FUNCTION_BLOCK PID_FLAG_STATE_ACCESS (* Experimental read-only state interface; original PID arithmetic unchanged; native validation pending *)
  (* Standard: 61499-2 *)
  (* Version 0.1, 2026-10-20, Guilherme *)
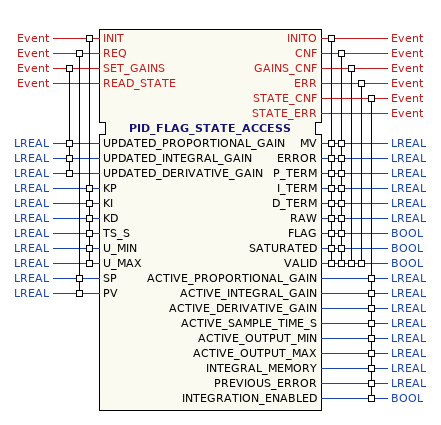
  EVENT_INPUT
    INIT WITH KP, KI, KD, TS_S, U_MIN, U_MAX;
    REQ WITH SP, PV;
    SET_GAINS WITH UPDATED_PROPORTIONAL_GAIN, UPDATED_INTEGRAL_GAIN, UPDATED_DERIVATIVE_GAIN;
    READ_STATE;
  END_EVENT
  EVENT_OUTPUT
    INITO WITH MV, ERROR, P_TERM, I_TERM, D_TERM, RAW, FLAG, SATURATED, VALID;
    CNF WITH MV, ERROR, P_TERM, I_TERM, D_TERM, RAW, FLAG, SATURATED, VALID;
    GAINS_CNF WITH VALID;
    ERR WITH VALID;
    STATE_CNF WITH ACTIVE_PROPORTIONAL_GAIN, ACTIVE_INTEGRAL_GAIN, ACTIVE_DERIVATIVE_GAIN, ACTIVE_SAMPLE_TIME_S, ACTIVE_OUTPUT_MIN, ACTIVE_OUTPUT_MAX, INTEGRAL_MEMORY, PREVIOUS_ERROR, INTEGRATION_ENABLED;
    STATE_ERR;
  END_EVENT
  VAR_INPUT
    UPDATED_PROPORTIONAL_GAIN : LREAL;
    UPDATED_INTEGRAL_GAIN : LREAL;
    UPDATED_DERIVATIVE_GAIN : LREAL;
    KP : LREAL;
    KI : LREAL;
    KD : LREAL;
    TS_S : LREAL;
    U_MIN : LREAL;
    U_MAX : LREAL;
    SP : LREAL;
    PV : LREAL;
  END_VAR
  VAR_OUTPUT
    MV : LREAL;
    ERROR : LREAL;
    P_TERM : LREAL;
    I_TERM : LREAL;
    D_TERM : LREAL;
    RAW : LREAL;
    FLAG : BOOL;
    SATURATED : BOOL;
    VALID : BOOL;
    ACTIVE_PROPORTIONAL_GAIN : LREAL;
    ACTIVE_INTEGRAL_GAIN : LREAL;
    ACTIVE_DERIVATIVE_GAIN : LREAL;
    ACTIVE_SAMPLE_TIME_S : LREAL;
    ACTIVE_OUTPUT_MIN : LREAL;
    ACTIVE_OUTPUT_MAX : LREAL;
    INTEGRAL_MEMORY : LREAL;
    PREVIOUS_ERROR : LREAL;
    INTEGRATION_ENABLED : BOOL;
  END_VAR
  VAR
    KP_ACTIVE : LREAL;
    KI_ACTIVE : LREAL;
    KD_ACTIVE : LREAL;
    TS_ACTIVE : LREAL;
    LOW : LREAL;
    HIGH : LREAL;
    I_MEMORY : LREAL;
    E_PREV : LREAL;
    E_NEXT : LREAL;
    I_NEXT : LREAL;
    D_NEXT : LREAL;
    P_NEXT : LREAL;
    IT_NEXT : LREAL;
    DT_NEXT : LREAL;
    RAW_NEXT : LREAL;
  END_VAR
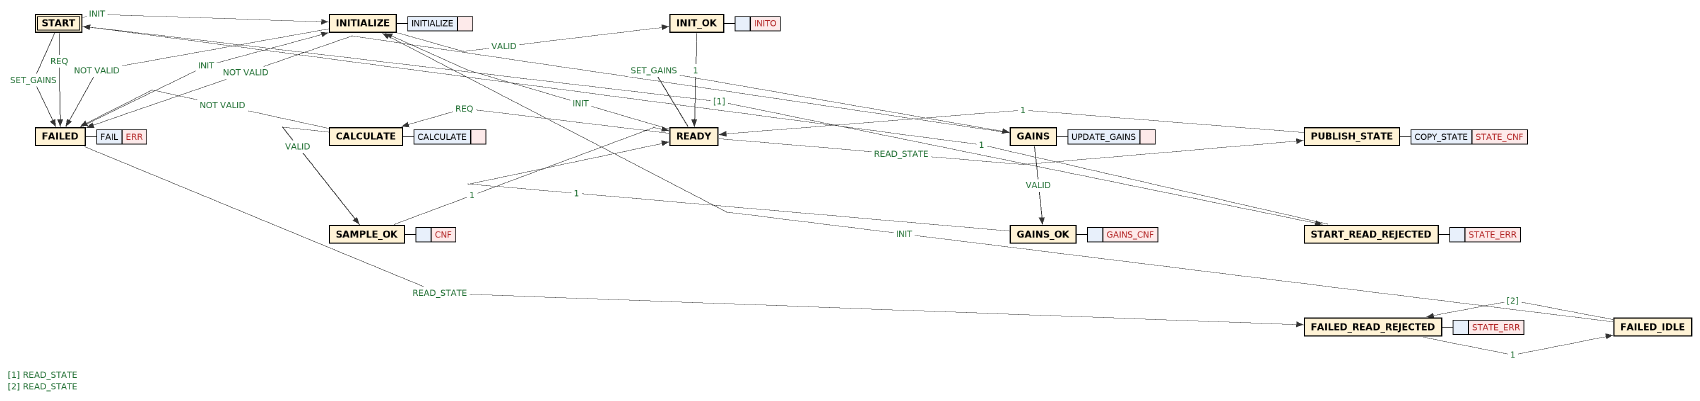
  EC_STATES
    START;
    FAILED_READ_REJECTED : -> STATE_ERR;
    START_READ_REJECTED : -> STATE_ERR;
    PUBLISH_STATE : COPY_STATE -> STATE_CNF;
    INITIALIZE : INITIALIZE;
    INIT_OK : -> INITO;
    READY;
    CALCULATE : CALCULATE;
    SAMPLE_OK : -> CNF;
    GAINS : UPDATE_GAINS;
    GAINS_OK : -> GAINS_CNF;
    FAILED : FAIL -> ERR;
    FAILED_IDLE;
  END_STATES
  EC_TRANSITIONS
    START TO INITIALIZE := INIT;
    START TO FAILED := REQ;
    START TO FAILED := SET_GAINS;
    INITIALIZE TO INIT_OK := VALID;
    INITIALIZE TO FAILED := NOT VALID;
    INIT_OK TO READY := 1;
    READY TO INITIALIZE := INIT;
    READY TO GAINS := SET_GAINS;
    READY TO CALCULATE := REQ;
    CALCULATE TO SAMPLE_OK := VALID;
    CALCULATE TO FAILED := NOT VALID;
    SAMPLE_OK TO READY := 1;
    GAINS TO GAINS_OK := VALID;
    GAINS TO FAILED := NOT VALID;
    GAINS_OK TO READY := 1;
    FAILED TO INITIALIZE := INIT;
    START TO START_READ_REJECTED := READ_STATE;
    START_READ_REJECTED TO START := 1;
    FAILED TO FAILED_READ_REJECTED := READ_STATE;
    FAILED_READ_REJECTED TO FAILED_IDLE := 1;
    FAILED_IDLE TO INITIALIZE := INIT;
    FAILED_IDLE TO FAILED_READ_REJECTED := READ_STATE;
    READY TO PUBLISH_STATE := READ_STATE;
    PUBLISH_STATE TO READY := 1;
  END_TRANSITIONS
  ALGORITHM INITIALIZE IN ST:
VALID := (KP >= -1.0E+100) AND (KP <= 1.0E+100) AND (KI >= -1.0E+100) AND (KI <= 1.0E+100) AND (KD >= -1.0E+100) AND (KD <= 1.0E+100) AND (TS_S >= -1.0E+100) AND (TS_S <= 1.0E+100) AND (U_MIN >= -1.0E+100) AND (U_MIN <= 1.0E+100) AND (U_MAX >= -1.0E+100) AND (U_MAX <= 1.0E+100) AND (TS_S > 0.0) AND (U_MIN < U_MAX);
IF VALID THEN
    KP_ACTIVE := KP;
    KI_ACTIVE := KI;
    KD_ACTIVE := KD;
    TS_ACTIVE := TS_S;
    LOW := U_MIN;
    HIGH := U_MAX;
    I_MEMORY := 0.0;
    E_PREV := 0.0;
    FLAG := TRUE;
    MV := 0.0;
    RAW := 0.0;
    ERROR := 0.0;
    P_TERM := 0.0;
    I_TERM := 0.0;
    D_TERM := 0.0;
    SATURATED := FALSE;
END_IF;
  END_ALGORITHM
  ALGORITHM CALCULATE IN ST:
VALID := (SP >= -1.0E+100) AND (SP <= 1.0E+100) AND (PV >= -1.0E+100) AND (PV <= 1.0E+100);
IF VALID THEN
    E_NEXT := SP - PV;
    I_NEXT := I_MEMORY;
    IF FLAG THEN
        I_NEXT := I_MEMORY + (TS_ACTIVE / 2.0) * (E_NEXT + E_PREV);
    END_IF;
    D_NEXT := (E_NEXT - E_PREV) / TS_ACTIVE;
    P_NEXT := KP_ACTIVE * E_NEXT;
    IT_NEXT := KI_ACTIVE * I_NEXT;
    DT_NEXT := KD_ACTIVE * D_NEXT;
    RAW_NEXT := P_NEXT + IT_NEXT + DT_NEXT;
    VALID := (E_NEXT >= -1.0E+100) AND (E_NEXT <= 1.0E+100) AND (I_NEXT >= -1.0E+100) AND (I_NEXT <= 1.0E+100) AND (D_NEXT >= -1.0E+100) AND (D_NEXT <= 1.0E+100) AND (P_NEXT >= -1.0E+100) AND (P_NEXT <= 1.0E+100) AND (IT_NEXT >= -1.0E+100) AND (IT_NEXT <= 1.0E+100) AND (DT_NEXT >= -1.0E+100) AND (DT_NEXT <= 1.0E+100) AND (RAW_NEXT >= -1.0E+100) AND (RAW_NEXT <= 1.0E+100);
    IF VALID THEN
        MV := RAW_NEXT;
        FLAG := TRUE;
        SATURATED := FALSE;
        IF RAW_NEXT > HIGH THEN
            MV := HIGH;
            FLAG := FALSE;
            SATURATED := TRUE;
        END_IF;
        IF RAW_NEXT < LOW THEN
            MV := LOW;
            FLAG := FALSE;
            SATURATED := TRUE;
        END_IF;
        I_MEMORY := I_NEXT;
        E_PREV := E_NEXT;
        ERROR := E_NEXT;
        P_TERM := P_NEXT;
        I_TERM := IT_NEXT;
        D_TERM := DT_NEXT;
        RAW := RAW_NEXT;
    END_IF;
END_IF;
  END_ALGORITHM
  ALGORITHM UPDATE_GAINS IN ST:
VALID := (UPDATED_PROPORTIONAL_GAIN >= -1.0E+100) AND (UPDATED_PROPORTIONAL_GAIN <= 1.0E+100) AND (UPDATED_INTEGRAL_GAIN >= -1.0E+100) AND (UPDATED_INTEGRAL_GAIN <= 1.0E+100) AND (UPDATED_DERIVATIVE_GAIN >= -1.0E+100) AND (UPDATED_DERIVATIVE_GAIN <= 1.0E+100);
IF VALID THEN
    KP_ACTIVE := UPDATED_PROPORTIONAL_GAIN;
    KI_ACTIVE := UPDATED_INTEGRAL_GAIN;
    KD_ACTIVE := UPDATED_DERIVATIVE_GAIN;
END_IF;
  END_ALGORITHM
  ALGORITHM FAIL IN ST:
VALID := FALSE;
  END_ALGORITHM
  ALGORITHM COPY_STATE IN ST:
ACTIVE_PROPORTIONAL_GAIN := KP_ACTIVE;
ACTIVE_INTEGRAL_GAIN := KI_ACTIVE;
ACTIVE_DERIVATIVE_GAIN := KD_ACTIVE;
ACTIVE_SAMPLE_TIME_S := TS_ACTIVE;
ACTIVE_OUTPUT_MIN := LOW;
ACTIVE_OUTPUT_MAX := HIGH;
INTEGRAL_MEMORY := I_MEMORY;
PREVIOUS_ERROR := E_PREV;
INTEGRATION_ENABLED := FLAG;
  END_ALGORITHM
END_FUNCTION_BLOCK
